# EPICS substitutions: db/MonoDAQ/ecmcMonoDAQ-E-gMeter.substitutions
file "ecmc_analogInput-chX.template"{
  pattern {CH_ID, KEY,      sourceName, ESLO, EGU,  PREC}
          {01,    counter,  counter,    1,    "",   0   }
}

file "ecmc_analogInputFloat-chX.template"{
  pattern {CH_ID, KEY,          sourceName,     ESLO, EGU,    PREC}
          {01,    temperature,  temperature,    1,    "degC", 3   }
          {01,    X,            accelerometerX, 1,    "g",    6   }
          {01,    Y,            accelerometerY, 1,    "g",    6   }
          {01,    Z,            accelerometerZ, 1,    "g",    6   }
}
